(* IEC 61131-3 sources: plc-vscode/tests/st/all/rusty/libs/stdlib/iec61131-st, 25 files *)

(* ---- arithmetic_functions.st ---- *)
(* Definitions of arithmetic functions defined by the IEC61131-3 standard *)

{external}
VAR_GLOBAL
    PI_REAL : REAL;
    PI_LREAL : LREAL;
    FRAC_PI_2_REAL : REAL;
    FRAC_PI_2_LREAL : LREAL;
    FRAC_PI_4_REAL : REAL;
    FRAC_PI_4_LREAL : LREAL;
    E_REAL : REAL;
    E_LREAL : LREAL;
    INF_REAL: REAL;
    INF_LREAL: LREAL;
    NAN_REAL: REAL;
    NAN_LREAL: LREAL;
END_VAR

(********************
*
* This operator returns the value of adding up the operands.
* It overloads the variadic builtin implementation of ADD, which is implemented for ANY_NUM
*
*********************)
FUNCTION ADD < T1: ANY, T2: ANY >: T1
VAR_INPUT
    IN1: T1;
    IN2: T2...;
END_VAR
END_FUNCTION

(********************
*
* This operator produces the multiplication of the operands.
* It overloads the variadic builtin implementation of MUL, which is implemented for ANY_NUM
*
*********************)
FUNCTION MUL < T1: ANY, T2: ANY >: T1
VAR_INPUT
    IN1: T1;
    IN2: T2...;
END_VAR
END_FUNCTION

(* Calculates the square root of a given value *)
{external}
FUNCTION SQRT<T : ANY_REAL> : T
VAR_INPUT
    in : T;
END_VAR
END_FUNCTION

(** Logarithmic functions **)

(* Calculates the natural logarithm of the given value *)
{external}
FUNCTION LN<T : ANY_REAL> : T
VAR_INPUT
    in : T;
END_VAR
END_FUNCTION

(* Calculates the base 10 logarithm of the given value *)
{external}
FUNCTION LOG<T : ANY_REAL> : T
VAR_INPUT
    in : T;
END_VAR
END_FUNCTION

(* Calculates the natural exporenent of the given value *)
{external}
FUNCTION EXP<T : ANY_REAL> : T
VAR_INPUT
    in : T;
END_VAR
END_FUNCTION

(** Trigonometric functions **)

(* Calculates the sine of the given value in radiants *)
{external}
FUNCTION SIN<T : ANY_REAL> : T
VAR_INPUT
    rad : T;
END_VAR
END_FUNCTION

(* Calculates the cosine of the given value in radiants *)
{external}
FUNCTION COS<T : ANY_REAL> : T
VAR_INPUT
    rad : T;
END_VAR
END_FUNCTION

(* Calculates the tangent of the given value in radiants *)
{external}
FUNCTION TAN<T : ANY_REAL> : T
VAR_INPUT
    rad : T;
END_VAR
END_FUNCTION

(* Calculates the arc sine of the given value *)
{external}
FUNCTION ASIN<T : ANY_REAL> : T
VAR_INPUT
    in : T;
END_VAR
END_FUNCTION

(* Calculates the arc cosine of the given value *)
{external}
FUNCTION ACOS<T : ANY_REAL> : T
VAR_INPUT
    in : T;
END_VAR
END_FUNCTION

(* Calculates the arc tangent of the given value *)
{external}
FUNCTION ATAN<T : ANY_REAL> : T
VAR_INPUT
    in : T;
END_VAR
END_FUNCTION

(* Calculate the four quadrant arc tangent of the given values *)
{external}
FUNCTION ATAN2<T : ANY_REAL> : T
VAR_INPUT
    y : T;
    x : T;
END_VAR
END_FUNCTION

{external}
FUNCTION EXPT<T: ANY_REAL, U: ANY_NUM> : T
VAR_INPUT
    in1 : T;
    in2 : U;
END_VAR
END_FUNCTION

{external}
FUNCTION EXPT__REAL__DINT : REAL
VAR_INPUT
    in1 : REAL;
    in2 : DINT;
END_VAR
END_FUNCTION

{external}
FUNCTION EXPT__REAL__REAL : REAL
VAR_INPUT
    in1 : REAL;
    in2 : REAL;
END_VAR
END_FUNCTION

(* LREAL to REAL conversion will happen for the exponent
   This will produce the closest possible REAL value
   On overflow, infinity of the same sign as the input is produced *)
{external}
FUNCTION EXPT__REAL__LREAL : REAL
VAR_INPUT
    in1 : REAL;
    in2 : LREAL;
END_VAR
END_FUNCTION

{external}
FUNCTION EXPT__LREAL__DINT : LREAL
VAR_INPUT
    in1 : LREAL;
    in2 : DINT;
END_VAR
END_FUNCTION

{external}
FUNCTION EXPT__LREAL__REAL : LREAL
VAR_INPUT
    in1 : LREAL;
    in2 : REAL;
END_VAR
END_FUNCTION

{external}
FUNCTION EXPT__LREAL__LREAL : LREAL
VAR_INPUT
    in1 : LREAL;
    in2 : LREAL;
END_VAR
END_FUNCTION

FUNCTION EXPT__REAL__USINT : REAL
VAR_INPUT
    in1 : REAL;
    in2 : USINT;
END_VAR
    EXPT__REAL__USINT := EXPT__REAL__DINT(in1, in2);
END_FUNCTION

FUNCTION EXPT__REAL__UINT : REAL
VAR_INPUT
    in1 : REAL;
    in2 : UINT;
END_VAR
    EXPT__REAL__UINT := EXPT__REAL__DINT(in1, in2);
END_FUNCTION

FUNCTION EXPT__REAL__UDINT : REAL
VAR_INPUT
    in1 : REAL;
    in2 : UDINT;
END_VAR
    EXPT__REAL__UDINT := EXPT__REAL__DINT(in1, in2);
END_FUNCTION

FUNCTION EXPT__REAL__ULINT : REAL
VAR_INPUT
    in1 : REAL;
    in2 : ULINT;
END_VAR
    EXPT__REAL__ULINT := EXPT__REAL__DINT(in1, in2);
END_FUNCTION

FUNCTION EXPT__REAL__SINT : REAL
VAR_INPUT
    in1 : REAL;
    in2 : SINT;
END_VAR
    EXPT__REAL__SINT := EXPT__REAL__DINT(in1, in2);
END_FUNCTION

FUNCTION EXPT__REAL__INT : REAL
VAR_INPUT
    in1 : REAL;
    in2 : INT;
END_VAR
    EXPT__REAL__INT := EXPT__REAL__DINT(in1, in2);
END_FUNCTION

FUNCTION EXPT__REAL__LINT : REAL
VAR_INPUT
    in1 : REAL;
    in2 : LINT;
END_VAR
    EXPT__REAL__LINT := EXPT__REAL__DINT(in1, in2);
END_FUNCTION

FUNCTION EXPT__LREAL__USINT : LREAL
VAR_INPUT
    in1 : LREAL;
    in2 : USINT;
END_VAR
    EXPT__LREAL__USINT := EXPT__LREAL__DINT(in1, in2);
END_FUNCTION

FUNCTION EXPT__LREAL__UINT : LREAL
VAR_INPUT
    in1 : LREAL;
    in2 : UINT;
END_VAR
    EXPT__LREAL__UINT := EXPT__LREAL__DINT(in1, in2);
END_FUNCTION

FUNCTION EXPT__LREAL__UDINT : LREAL
VAR_INPUT
    in1 : LREAL;
    in2 : UDINT;
END_VAR
    EXPT__LREAL__UDINT := EXPT__LREAL__DINT(in1, in2);
END_FUNCTION

FUNCTION EXPT__LREAL__ULINT : LREAL
VAR_INPUT
    in1 : LREAL;
    in2 : ULINT;
END_VAR
    EXPT__LREAL__ULINT := EXPT__LREAL__DINT(in1, in2);
END_FUNCTION

FUNCTION EXPT__LREAL__SINT : LREAL
VAR_INPUT
    in1 : LREAL;
    in2 : SINT;
END_VAR
    EXPT__LREAL__SINT := EXPT__LREAL__DINT(in1, in2);
END_FUNCTION

FUNCTION EXPT__LREAL__INT : LREAL
VAR_INPUT
    in1 : LREAL;
    in2 : INT;
END_VAR
    EXPT__LREAL__INT := EXPT__LREAL__DINT(in1, in2);
END_FUNCTION

FUNCTION EXPT__LREAL__LINT : LREAL
VAR_INPUT
    in1 : LREAL;
    in2 : LINT;
END_VAR
    EXPT__LREAL__LINT := EXPT__LREAL__DINT(in1, in2);
END_FUNCTION

(* ---- string_functions.st ---- *)
VAR_GLOBAL CONSTANT
    __STRING_LENGTH: DINT := 2048;
END_VAR

(* *****************************************************************************
Description: String character length
Input:
    - IN: A character string
Return: String length
***************************************************************************** *)
{external}
FUNCTION LEN < T: ANY_STRING >: DINT
VAR_INPUT {ref}
    IN: T;
END_VAR
END_FUNCTION

(* *****************************************************************************
Description: Left
Input:
    - IN: A character string
    - L: The length of the substring
Return: A substring consisting of the leftmost L characters of IN
***************************************************************************** *)
FUNCTION LEFT < T: ANY_STRING >: T
VAR_INPUT {ref}
    IN: T;
END_VAR
VAR_INPUT
    L: DINT;
END_VAR
END_FUNCTION

{external}
FUNCTION LEFT_EXT < T: ANY_STRING >: DINT
VAR_INPUT {ref}
    IN: T;
END_VAR
VAR_INPUT
    L: DINT;
END_VAR
VAR_IN_OUT
    OUT: T;
END_VAR
END_FUNCTION

FUNCTION LEFT__STRING: STRING[__STRING_LENGTH]
VAR_INPUT {ref}
    IN: STRING[__STRING_LENGTH];
END_VAR
VAR_INPUT
    L: DINT;
END_VAR
    LEFT_EXT(IN, L, LEFT__STRING);
END_FUNCTION

FUNCTION LEFT__WSTRING: WSTRING[__STRING_LENGTH]
VAR_INPUT {ref}
    IN: WSTRING[__STRING_LENGTH];
END_VAR
VAR_INPUT
    L: DINT;
END_VAR
    LEFT_EXT(IN, L, LEFT__WSTRING);
END_FUNCTION

{external}
FUNCTION LEFT_EXT__STRING: DINT
VAR_INPUT {ref}
    IN: STRING[__STRING_LENGTH];
END_VAR
VAR_INPUT
    L: DINT;
END_VAR
VAR_IN_OUT
    OUT: STRING[__STRING_LENGTH];
END_VAR
END_FUNCTION

{external}
FUNCTION LEFT_EXT__WSTRING: DINT
VAR_INPUT {ref}
    IN: WSTRING[__STRING_LENGTH];
END_VAR
VAR_INPUT
    L: DINT;
END_VAR
VAR_IN_OUT
    OUT: WSTRING[__STRING_LENGTH];
END_VAR
END_FUNCTION

(* *****************************************************************************
Description: Right
Input:
    - IN: A character string
    - L: The length of the substring
Return: A substring consisting of the rightmost L characters of IN
***************************************************************************** *)
FUNCTION RIGHT < T: ANY_STRING >: T
VAR_INPUT {ref}
    IN: T;
END_VAR
VAR_INPUT
    L: DINT;
END_VAR
END_FUNCTION

{external}
FUNCTION RIGHT_EXT < T: ANY_STRING >: DINT
VAR_INPUT {ref}
    IN: T;
END_VAR
VAR_INPUT
    L: DINT;
END_VAR
VAR_IN_OUT
    OUT: T;
END_VAR
END_FUNCTION

FUNCTION RIGHT__STRING: STRING[__STRING_LENGTH]
VAR_INPUT {ref}
    IN: STRING[__STRING_LENGTH];
END_VAR
VAR_INPUT
    L: DINT;
END_VAR
    RIGHT_EXT(IN, L, RIGHT__STRING);
END_FUNCTION

FUNCTION RIGHT__WSTRING: WSTRING[__STRING_LENGTH]
VAR_INPUT {ref}
    IN: WSTRING[__STRING_LENGTH];
END_VAR
VAR_INPUT
    L: DINT;
END_VAR
    RIGHT_EXT(IN, L, RIGHT__WSTRING);
END_FUNCTION

{external}
FUNCTION RIGHT_EXT__STRING: DINT
VAR_INPUT {ref}
    IN: STRING[__STRING_LENGTH];
END_VAR
VAR_INPUT
    L: DINT;
END_VAR
VAR_IN_OUT
    OUT: STRING[__STRING_LENGTH];
END_VAR
END_FUNCTION

{external}
FUNCTION RIGHT_EXT__WSTRING: DINT
VAR_INPUT {ref}
    IN: WSTRING[__STRING_LENGTH];
END_VAR
VAR_INPUT
    L: DINT;
END_VAR
VAR_IN_OUT
    OUT: WSTRING[__STRING_LENGTH];
END_VAR
END_FUNCTION

(* *****************************************************************************
Description: Middle
Input:
    - IN: A character string
    - L: The length of the substring
    - P: The starting index position
Return:
    A substring that contains L characters starting
    from position P in a string.
***************************************************************************** *)
FUNCTION MID < T: ANY_STRING >: T
VAR_INPUT {ref}
    IN: T;
END_VAR
VAR_INPUT
    L: DINT;
    P: DINT;
END_VAR
END_FUNCTION

{external}
FUNCTION MID_EXT < T: ANY_STRING >: DINT
VAR_INPUT {ref}
    IN: T;
END_VAR
VAR_INPUT
    L: DINT;
    P: DINT;
END_VAR
VAR_IN_OUT
    OUT: T;
END_VAR
END_FUNCTION

FUNCTION MID__STRING: STRING[__STRING_LENGTH]
VAR_INPUT {ref}
    IN: STRING[__STRING_LENGTH];
END_VAR
VAR_INPUT
    L: DINT;
    P: DINT;
END_VAR
    MID_EXT(IN, L, P, MID__STRING);
END_FUNCTION

FUNCTION MID__WSTRING: WSTRING[__STRING_LENGTH]
VAR_INPUT {ref}
    IN: WSTRING[__STRING_LENGTH];
END_VAR
VAR_INPUT
    L: DINT;
    P: DINT;
END_VAR
    MID_EXT(IN, L, P, MID__WSTRING);
END_FUNCTION

{external}
FUNCTION MID_EXT__STRING: DINT
VAR_INPUT {ref}
    IN: STRING[__STRING_LENGTH];
END_VAR
VAR_INPUT
    L: DINT;
    P: DINT;
END_VAR
VAR_IN_OUT
    OUT: STRING[__STRING_LENGTH];
END_VAR
END_FUNCTION

{external}
FUNCTION MID_EXT__WSTRING: DINT
VAR_INPUT {ref}
    IN: WSTRING[__STRING_LENGTH];
END_VAR
VAR_INPUT
    L: DINT;
    P: DINT;
END_VAR
VAR_IN_OUT
    OUT: WSTRING[__STRING_LENGTH];
END_VAR
END_FUNCTION

(* *****************************************************************************
Description: Extensible concatenation
Input:
    - IN: Two or more comma-separated strings
Return:
    A string combining all given input strings in the same order
    as the given string parameters.
***************************************************************************** *)
{external}
FUNCTION CONCAT__STRING: STRING[2048]
VAR_INPUT {ref}
    args: {sized} STRING...;
END_VAR
END_FUNCTION

{external}
FUNCTION CONCAT__WSTRING: WSTRING[2048]
VAR_INPUT {ref}
    args: {sized} WSTRING...;
END_VAR
END_FUNCTION

FUNCTION CONCAT < T: ANY_STRING >: T
VAR_INPUT {ref}
    args: {sized} T...;
END_VAR
END_FUNCTION

{external}
FUNCTION CONCAT_EXT < T: ANY_STRING >: DINT
VAR_IN_OUT
    OUT: T;
END_VAR
VAR_INPUT {ref}
    args: {sized} T...;
END_VAR
END_FUNCTION

(* *****************************************************************************
Description: Insert
Input:
    IN1: The string to insert into
    IN2: The string to insert
    P: The position at which to insert
Return:
    A string consisting of IN2 inserted at position P into string IN1
***************************************************************************** *)
FUNCTION INSERT < T: ANY_STRING >: T
VAR_INPUT {ref}
    IN1: T;
    IN2: T;
END_VAR
VAR_INPUT
    P: DINT;
END_VAR
END_FUNCTION

{external}
FUNCTION INSERT_EXT < T: ANY_STRING >: DINT
VAR_INPUT {ref}
    IN1: T;
    IN2: T;
END_VAR
VAR_INPUT
    P: DINT;
END_VAR
VAR_IN_OUT
    OUT: T;
END_VAR
END_FUNCTION

FUNCTION INSERT__STRING: STRING[__STRING_LENGTH]
VAR_INPUT {ref}
    IN1: STRING[__STRING_LENGTH];
    IN2: STRING[__STRING_LENGTH];
END_VAR
VAR_INPUT
    P: DINT;
END_VAR
    INSERT_EXT(IN1, IN2, P, INSERT__STRING);
END_FUNCTION

FUNCTION INSERT__WSTRING: WSTRING[__STRING_LENGTH]
VAR_INPUT {ref}
    IN1: WSTRING[__STRING_LENGTH];
    IN2: WSTRING[__STRING_LENGTH];
END_VAR
VAR_INPUT
    P: DINT;
END_VAR
    INSERT_EXT(IN1, IN2, P, INSERT__WSTRING);
END_FUNCTION

{external}
FUNCTION INSERT_EXT__STRING: DINT
VAR_INPUT {ref}
    IN1: STRING[__STRING_LENGTH];
    IN2: STRING[__STRING_LENGTH];
END_VAR
VAR_INPUT
    P: DINT;
END_VAR
VAR_IN_OUT
    OUT: STRING[__STRING_LENGTH];
END_VAR
END_FUNCTION

{external}
FUNCTION INSERT_EXT__WSTRING: DINT
VAR_INPUT {ref}
    IN1: WSTRING[__STRING_LENGTH];
    IN2: WSTRING[__STRING_LENGTH];
END_VAR
VAR_INPUT
    P: DINT;
END_VAR
VAR_IN_OUT
    OUT: WSTRING[__STRING_LENGTH];
END_VAR
END_FUNCTION

(* *****************************************************************************
Description: Delete
Input:
    IN: The string to delete characters from
    L: The amount of characters to delete
    P: The position at which to start deleting
Return: A new string with L characters deleted from P onwards
***************************************************************************** *)
FUNCTION DELETE < T: ANY_STRING >: T
VAR_INPUT {ref}
    IN: T;
END_VAR
VAR_INPUT
    L: DINT;
    P: DINT;
END_VAR
END_FUNCTION

{external}
FUNCTION DELETE_EXT < T: ANY_STRING >: DINT
VAR_INPUT {ref}
    IN: T;
END_VAR
VAR_INPUT
    L: DINT;
    P: DINT;
END_VAR
VAR_IN_OUT
    OUT: T;
END_VAR
END_FUNCTION

FUNCTION DELETE__STRING: STRING[__STRING_LENGTH]
VAR_INPUT {ref}
    IN: STRING[__STRING_LENGTH];
END_VAR
VAR_INPUT
    L: DINT;
    P: DINT;
END_VAR
    DELETE_EXT(IN, L, P, DELETE__STRING);
END_FUNCTION

FUNCTION DELETE__WSTRING: WSTRING[__STRING_LENGTH]
VAR_INPUT {ref}
    IN: WSTRING[__STRING_LENGTH];
END_VAR
VAR_INPUT
    L: DINT;
    P: DINT;
END_VAR
    DELETE_EXT(IN, L, P, DELETE__WSTRING);
END_FUNCTION

{external}
FUNCTION DELETE_EXT__STRING: DINT
VAR_INPUT {ref}
    IN: STRING[__STRING_LENGTH];
END_VAR
VAR_INPUT
    L: DINT;
    P: DINT;
END_VAR
VAR_IN_OUT
    OUT: STRING[__STRING_LENGTH];
END_VAR
END_FUNCTION

{external}
FUNCTION DELETE_EXT__WSTRING: DINT
VAR_INPUT {ref}
    IN: WSTRING[__STRING_LENGTH];
END_VAR
VAR_INPUT
    L: DINT;
    P: DINT;
END_VAR
VAR_IN_OUT
    OUT: WSTRING[__STRING_LENGTH];
END_VAR
END_FUNCTION
(* *****************************************************************************
Description: Replace
Input:
    IN1: The string to replace characters from
    IN2: The replacement string to be inserted
    L: The amount of characters to delete
    P: The position at which to start deleting
Return: A new string which has L characters replaced by IN2 from position P onwards
***************************************************************************** *)
FUNCTION REPLACE < T: ANY_STRING >: T
VAR_INPUT {ref}
    IN1: T;
    IN2: T;
END_VAR
VAR_INPUT
    L: DINT;
    P: DINT;
END_VAR
END_FUNCTION

{external}
FUNCTION REPLACE_EXT < T: ANY_STRING >: DINT
VAR_INPUT {ref}
    IN1: T;
    IN2: T;
END_VAR
VAR_INPUT
    L: DINT;
    P: DINT;
END_VAR
VAR_IN_OUT
    OUT: T;
END_VAR
END_FUNCTION

FUNCTION REPLACE__STRING: STRING[__STRING_LENGTH]
VAR_INPUT {ref}
    IN1: STRING[__STRING_LENGTH];
    IN2: STRING[__STRING_LENGTH];
END_VAR
VAR_INPUT
    L: DINT;
    P: DINT;
END_VAR
    REPLACE_EXT(IN1, IN2, L, P, REPLACE__STRING);
END_FUNCTION

FUNCTION REPLACE__WSTRING: WSTRING[__STRING_LENGTH]
VAR_INPUT {ref}
    IN1: WSTRING[__STRING_LENGTH];
    IN2: WSTRING[__STRING_LENGTH];
END_VAR
VAR_INPUT
    L: DINT;
    P: DINT;
END_VAR
    REPLACE_EXT(IN1, IN2, L, P, REPLACE__WSTRING);
END_FUNCTION

{external}
FUNCTION REPLACE_EXT__STRING: DINT
VAR_INPUT {ref}
    IN1: STRING[__STRING_LENGTH];
    IN2: STRING[__STRING_LENGTH];
END_VAR
VAR_INPUT
    L: DINT;
    P: DINT;
END_VAR
VAR_IN_OUT
    OUT: STRING[__STRING_LENGTH];
END_VAR
END_FUNCTION

{external}
FUNCTION REPLACE_EXT__WSTRING: DINT
VAR_INPUT {ref}
    IN1: WSTRING[__STRING_LENGTH];
    IN2: WSTRING[__STRING_LENGTH];
END_VAR
VAR_INPUT
    L: DINT;
    P: DINT;
END_VAR
VAR_IN_OUT
    OUT: WSTRING[__STRING_LENGTH];
END_VAR
END_FUNCTION

(* *****************************************************************************
Description: Find
Input:
    IN1: The string in which to search in
    IN2: The substring to search for
Return: The character index of the first match. 0 if there are no matches.
***************************************************************************** *)
{external}
FUNCTION FIND < T: ANY_STRING >: DINT
VAR_INPUT {ref}
    IN1: T;
    IN2: T;
END_VAR
END_FUNCTION

(* *****************************************************************************
Description: Decreasing sequence
Input: The strings to compare, in order. ((IN1>IN2) & (IN2>IN3) & .. & (INn-1>INn))
Return:
    TRUE if codepoints are in decreasing order (alphabetical order: ZYX > YXW > XWV ..)
    FALSE otherwise
***************************************************************************** *)
// passing strings by ref causes an error/warning. code still compiles and works correctly
FUNCTION STRING_GREATER: BOOL
VAR_INPUT
    a, b: STRING;
END_VAR
    STRING_GREATER := __STRING_GREATER(a, b);
END_FUNCTION

FUNCTION WSTRING_GREATER: BOOL
VAR_INPUT
    a, b: WSTRING;
END_VAR
    WSTRING_GREATER := __WSTRING_GREATER(a, b);
END_FUNCTION

(* *****************************************************************************
Description: Equality
Input: The strings to compare, in order. ((IN1=IN2) & (IN2=IN3) & .. & (INn-1=INn))
Return:
    TRUE if codepoints are equal to each other
    FALSE otherwise.
***************************************************************************** *)
FUNCTION STRING_EQUAL: BOOL
VAR_INPUT
    a, b: STRING;
END_VAR
    STRING_EQUAL := __STRING_EQUAL(a, b);
END_FUNCTION

FUNCTION WSTRING_EQUAL: BOOL
VAR_INPUT
    a, b: WSTRING;
END_VAR
    WSTRING_EQUAL := __WSTRING_EQUAL(a, b);
END_FUNCTION

(* *****************************************************************************
Description: Increasing sequence
Input: The strings to compare, in order. ((IN1<IN2) & (IN2<IN3) & .. & (INn-1<INn))
Return:
    TRUE if codepoints are in increasing order (alphabetical order: ABC < BCD < CDE ..)
    FALSE otherwise
***************************************************************************** *)
FUNCTION STRING_LESS: BOOL
VAR_INPUT
    a, b: STRING;
END_VAR
    STRING_LESS := __STRING_LESS(a, b);
END_FUNCTION

FUNCTION WSTRING_LESS: BOOL
VAR_INPUT
    a, b: WSTRING;
END_VAR
    WSTRING_LESS := __WSTRING_LESS(a, b);
END_FUNCTION

// internal functions
{external}
FUNCTION __STRING_GREATER: BOOL
VAR_INPUT {ref}
    IN: {sized} STRING...;
END_VAR
END_FUNCTION

{external}
FUNCTION __STRING_EQUAL: BOOL
VAR_INPUT {ref}
    IN: {sized} STRING...;
END_VAR
END_FUNCTION

{external}
FUNCTION __STRING_LESS: BOOL
VAR_INPUT {ref}
    IN: {sized} STRING...;
END_VAR
END_FUNCTION

{external}
FUNCTION __WSTRING_GREATER: BOOL
VAR_INPUT {ref}
    IN: {sized} WSTRING...;
END_VAR
END_FUNCTION

{external}
FUNCTION __WSTRING_EQUAL: BOOL
VAR_INPUT {ref}
    IN: {sized} WSTRING...;
END_VAR
END_FUNCTION

{external}
FUNCTION __WSTRING_LESS: BOOL
VAR_INPUT {ref}
    IN: {sized} WSTRING...;
END_VAR
END_FUNCTION

(* ---- bit_conversion.st ---- *)
(********************
*
* Converts LWORD to DWORD
*
*********************)
FUNCTION LWORD_TO_DWORD : DWORD
VAR_INPUT
    in : LWORD;
END_VAR
    LWORD_TO_DWORD := in;
END_FUNCTION

(********************
*
* Converts LWORD to WORD
*
*********************)
FUNCTION LWORD_TO_WORD : WORD
VAR_INPUT
    in : LWORD;
END_VAR
    LWORD_TO_WORD := in;
END_FUNCTION

(********************
*
* Converts LWORD to BYTE
*
*********************)
FUNCTION LWORD_TO_BYTE : BYTE
VAR_INPUT
    in : LWORD;
END_VAR
    LWORD_TO_BYTE := in;
END_FUNCTION

(********************
*
* Converts LWORD to BOOL
*
*********************)
FUNCTION LWORD_TO_BOOL : BOOL
VAR_INPUT
    in : LWORD;
END_VAR
    LWORD_TO_BOOL := in.0;
END_FUNCTION

(********************
*
* Converts DWORD to LWORD
*
*********************)
FUNCTION DWORD_TO_LWORD : LWORD
VAR_INPUT
    in : DWORD;
END_VAR
    DWORD_TO_LWORD := in;
END_FUNCTION

(********************
*
* Converts DWORD to WORD
*
*********************)
FUNCTION DWORD_TO_WORD : WORD
VAR_INPUT
    in : DWORD;
END_VAR
    DWORD_TO_WORD := in;
END_FUNCTION

(********************
*
* Converts DWORD to BYTE
*
*********************)
FUNCTION DWORD_TO_BYTE : BYTE
VAR_INPUT
    in : DWORD;
END_VAR
    DWORD_TO_BYTE := in;
END_FUNCTION

(********************
*
* Converts DWORD to BOOL
*
*********************)
FUNCTION DWORD_TO_BOOL : BOOL
VAR_INPUT
    in : DWORD;
END_VAR
    DWORD_TO_BOOL := in.0;
END_FUNCTION

(********************
*
* Converts WORD to LWORD
*
*********************)
FUNCTION WORD_TO_LWORD : LWORD
VAR_INPUT
    in : WORD;
END_VAR
    WORD_TO_LWORD := in;
END_FUNCTION

(********************
*
* Converts WORD to DWORD
*
*********************)
FUNCTION WORD_TO_DWORD : DWORD
VAR_INPUT
    in : WORD;
END_VAR
    WORD_TO_DWORD := in;
END_FUNCTION

(********************
*
* Converts WORD to BYTE
*
*********************)
FUNCTION WORD_TO_BYTE : BYTE
VAR_INPUT
    in : WORD;
END_VAR
    WORD_TO_BYTE := in;
END_FUNCTION

(********************
*
* Converts WORD to BOOL
*
*********************)
FUNCTION WORD_TO_BOOL : BOOL
VAR_INPUT
    in : WORD;
END_VAR
    WORD_TO_BOOL := in.0;
END_FUNCTION

(********************
*
* Converts BYTE to LWORD
*
*********************)
FUNCTION BYTE_TO_LWORD : LWORD
VAR_INPUT
    in : BYTE;
END_VAR
    BYTE_TO_LWORD := in;
END_FUNCTION

(********************
*
* Converts BYTE to DWORD
*
*********************)
FUNCTION BYTE_TO_DWORD : DWORD
VAR_INPUT
    in : BYTE;
END_VAR
    BYTE_TO_DWORD := in;
END_FUNCTION

(********************
*
* Converts BYTE to WORD
*
*********************)
FUNCTION BYTE_TO_WORD : WORD
VAR_INPUT
    in : BYTE;
END_VAR
    BYTE_TO_WORD := in;
END_FUNCTION

(********************
*
* Converts BYTE to BOOL
*
*********************)
FUNCTION BYTE_TO_BOOL : BOOL
VAR_INPUT
    in : BYTE;
END_VAR
    BYTE_TO_BOOL := in.0;
END_FUNCTION

(********************
*
* Converts BYTE to CHAR
*
*********************)
FUNCTION BYTE_TO_CHAR : CHAR
VAR_INPUT
    in : BYTE;
END_VAR
VAR
    ptr : REF_TO CHAR;
END_VAR
    ptr := REF(in);
    BYTE_TO_CHAR := ptr^;
END_FUNCTION

(********************
*
* Converts BOOL to LWORD
*
*********************)
FUNCTION BOOL_TO_LWORD : LWORD
VAR_INPUT
    in : BOOL;
END_VAR
    IF in <> 0 THEN
        BOOL_TO_LWORD := 1;
    ELSE
        BOOL_TO_LWORD := 0;
    END_IF;
END_FUNCTION

(********************
*
* Converts BOOL to DWORD
*
*********************)
FUNCTION BOOL_TO_DWORD : DWORD
VAR_INPUT
    in : BOOL;
END_VAR
    IF in <> 0 THEN
        BOOL_TO_DWORD := 1;
    ELSE
        BOOL_TO_DWORD := 0;
    END_IF;
END_FUNCTION

(********************
*
* Converts BOOL to WORD
*
*********************)
FUNCTION BOOL_TO_WORD : WORD
VAR_INPUT
    in : BOOL;
END_VAR
    IF in <> 0 THEN
        BOOL_TO_WORD := 1;
    ELSE
        BOOL_TO_WORD := 0;
    END_IF;
END_FUNCTION

(********************
*
* Converts BOOL to BYTE
*
*********************)
FUNCTION BOOL_TO_BYTE : BYTE
VAR_INPUT
    in : BOOL;
END_VAR
    IF in <> 0 THEN
        BOOL_TO_BYTE := 1;
    ELSE
        BOOL_TO_BYTE := 0;
    END_IF;
END_FUNCTION

(********************
*
* Converts CHAR to BYTE
*
*********************)
FUNCTION CHAR_TO_BYTE : BYTE
VAR_INPUT
    in : CHAR;
END_VAR
VAR
    ptr : REF_TO BYTE;
END_VAR
    ptr := REF(in);
    CHAR_TO_BYTE := ptr^;
END_FUNCTION

(********************
*
* Converts WCHAR to BYTE
*
*********************)
FUNCTION WCHAR_TO_BYTE : BYTE
VAR_INPUT
    in : WCHAR;
END_VAR
VAR
    ptr : REF_TO BYTE;
END_VAR
    ptr := REF(in);
    WCHAR_TO_BYTE := ptr^;
END_FUNCTION

(********************
*
* Converts CHAR to WORD
*
*********************)
FUNCTION CHAR_TO_WORD : WORD
VAR_INPUT
    in : CHAR;
END_VAR
    CHAR_TO_WORD := CHAR_TO_BYTE(in);
END_FUNCTION

(********************
*
* Converts CHAR to DWORD
*
*********************)
FUNCTION CHAR_TO_DWORD : DWORD
VAR_INPUT
    in : CHAR;
END_VAR
    CHAR_TO_DWORD := CHAR_TO_BYTE(in);
END_FUNCTION

(********************
*
* Converts CHAR to LWORD
*
*********************)
FUNCTION CHAR_TO_LWORD : LWORD
VAR_INPUT
    in : CHAR;
END_VAR
    CHAR_TO_LWORD := CHAR_TO_BYTE(in);
END_FUNCTION

(********************
*
* Converts WCHAR to WORD
*
*********************)
FUNCTION WCHAR_TO_WORD : WORD
VAR_INPUT
    in : WCHAR;
END_VAR
VAR
    ptr : REF_TO WORD;
END_VAR
    ptr := REF(in);
    WCHAR_TO_WORD := ptr^;
END_FUNCTION

(********************
*
* Converts WCHAR to DWORD
*
*********************)
FUNCTION WCHAR_TO_DWORD : DWORD
VAR_INPUT
    in : WCHAR;
END_VAR
    WCHAR_TO_DWORD := WCHAR_TO_WORD(in);
END_FUNCTION

(********************
*
* Converts WCHAR to LWORD
*
*********************)
FUNCTION WCHAR_TO_LWORD : LWORD
VAR_INPUT
    in : WCHAR;
END_VAR
    WCHAR_TO_LWORD := WCHAR_TO_WORD(in);
END_FUNCTION

(* ---- bit_num_conversion.st ---- *)
(********************
*
* Converts LWORD to LREAL
*
*********************)
{external}
FUNCTION LWORD_TO_LREAL : LREAL
VAR_INPUT
    in : LWORD;
END_VAR
END_FUNCTION

(********************
*
* Converts LWORD to LINT
*
*********************)
FUNCTION LWORD_TO_LINT : LINT
VAR_INPUT
    in : LWORD;
END_VAR
    LWORD_TO_LINT := in;
END_FUNCTION

(********************
*
* Converts LWORD to DINT
*
*********************)
FUNCTION LWORD_TO_DINT : DINT
VAR_INPUT
    in : LWORD;
END_VAR
    LWORD_TO_DINT := in;
END_FUNCTION

(********************
*
* Converts LWORD to INT
*
*********************)
FUNCTION LWORD_TO_INT : INT
VAR_INPUT
    in : LWORD;
END_VAR
    LWORD_TO_INT := in;
END_FUNCTION

(********************
*
* Converts LWORD to SINT
*
*********************)
FUNCTION LWORD_TO_SINT : SINT
VAR_INPUT
    in : LWORD;
END_VAR
    LWORD_TO_SINT := in;
END_FUNCTION

(********************
*
* Converts LWORD to ULINT
*
*********************)
FUNCTION LWORD_TO_ULINT : ULINT
VAR_INPUT
    in : LWORD;
END_VAR
    LWORD_TO_ULINT := in;
END_FUNCTION

(********************
*
* Converts LWORD to UDINT
*
*********************)
FUNCTION LWORD_TO_UDINT : UDINT
VAR_INPUT
    in : LWORD;
END_VAR
    LWORD_TO_UDINT := in;
END_FUNCTION

(********************
*
* Converts LWORD to UINT
*
*********************)
FUNCTION LWORD_TO_UINT : UINT
VAR_INPUT
    in : LWORD;
END_VAR
    LWORD_TO_UINT := in;
END_FUNCTION

(********************
*
* Converts LWORD to USINT
*
*********************)
FUNCTION LWORD_TO_USINT : USINT
VAR_INPUT
    in : LWORD;
END_VAR
    LWORD_TO_USINT := in;
END_FUNCTION

(********************
*
* Converts DWORD to REAL
*
*********************)
{external}
FUNCTION DWORD_TO_REAL : REAL
VAR_INPUT
    in : DWORD;
END_VAR
END_FUNCTION

(********************
*
* Converts DWORD to LINT
*
*********************)
FUNCTION DWORD_TO_LINT : LINT
VAR_INPUT
    in : DWORD;
END_VAR
    DWORD_TO_LINT := in;
END_FUNCTION

(********************
*
* Converts DWORD to DINT
*
*********************)
FUNCTION DWORD_TO_DINT : DINT
VAR_INPUT
    in : DWORD;
END_VAR
    DWORD_TO_DINT := in;
END_FUNCTION

(********************
*
* Converts DWORD to INT
*
*********************)
FUNCTION DWORD_TO_INT : INT
VAR_INPUT
    in : DWORD;
END_VAR
    DWORD_TO_INT := in;
END_FUNCTION

(********************
*
* Converts DWORD to SINT
*
*********************)
FUNCTION DWORD_TO_SINT : SINT
VAR_INPUT
    in : DWORD;
END_VAR
    DWORD_TO_SINT := in;
END_FUNCTION

(********************
*
* Converts DWORD to ULINT
*
*********************)
FUNCTION DWORD_TO_ULINT : ULINT
VAR_INPUT
    in : DWORD;
END_VAR
    DWORD_TO_ULINT := in;
END_FUNCTION

(********************
*
* Converts DWORD to UDINT
*
*********************)
FUNCTION DWORD_TO_UDINT : UDINT
VAR_INPUT
    in : DWORD;
END_VAR
    DWORD_TO_UDINT := in;
END_FUNCTION

(********************
*
* Converts DWORD to UINT
*
*********************)
FUNCTION DWORD_TO_UINT : UINT
VAR_INPUT
    in : DWORD;
END_VAR
    DWORD_TO_UINT := in;
END_FUNCTION

(********************
*
* Converts DWORD to USINT
*
*********************)
FUNCTION DWORD_TO_USINT : USINT
VAR_INPUT
    in : DWORD;
END_VAR
    DWORD_TO_USINT := in;
END_FUNCTION

(********************
*
* Converts WORD to LINT
*
*********************)
FUNCTION WORD_TO_LINT : LINT
VAR_INPUT
    in : WORD;
END_VAR
    WORD_TO_LINT := in;
END_FUNCTION

(********************
*
* Converts WORD to DINT
*
*********************)
FUNCTION WORD_TO_DINT : DINT
VAR_INPUT
    in : WORD;
END_VAR
    WORD_TO_DINT := in;
END_FUNCTION

(********************
*
* Converts WORD to INT
*
*********************)
FUNCTION WORD_TO_INT : INT
VAR_INPUT
    in : WORD;
END_VAR
    WORD_TO_INT := in;
END_FUNCTION

(********************
*
* Converts WORD to SINT
*
*********************)
FUNCTION WORD_TO_SINT : SINT
VAR_INPUT
    in : WORD;
END_VAR
    WORD_TO_SINT := in;
END_FUNCTION

(********************
*
* Converts WORD to ULINT
*
*********************)
FUNCTION WORD_TO_ULINT : ULINT
VAR_INPUT
    in : WORD;
END_VAR
    WORD_TO_ULINT := in;
END_FUNCTION

(********************
*
* Converts WORD to UDINT
*
*********************)
FUNCTION WORD_TO_UDINT : UDINT
VAR_INPUT
    in : WORD;
END_VAR
    WORD_TO_UDINT := in;
END_FUNCTION

(********************
*
* Converts WORD to UINT
*
*********************)
FUNCTION WORD_TO_UINT : UINT
VAR_INPUT
    in : WORD;
END_VAR
    WORD_TO_UINT := in;
END_FUNCTION

(********************
*
* Converts WORD to USINT
*
*********************)
FUNCTION WORD_TO_USINT : USINT
VAR_INPUT
    in : WORD;
END_VAR
    WORD_TO_USINT := in;
END_FUNCTION

(********************
*
* Converts BYTE to LINT
*
*********************)
FUNCTION BYTE_TO_LINT : LINT
VAR_INPUT
    in : BYTE;
END_VAR
    BYTE_TO_LINT := in;
END_FUNCTION

(********************
*
* Converts BYTE to DINT
*
*********************)
FUNCTION BYTE_TO_DINT : DINT
VAR_INPUT
    in : BYTE;
END_VAR
    BYTE_TO_DINT := in;
END_FUNCTION

(********************
*
* Converts BYTE to INT
*
*********************)
FUNCTION BYTE_TO_INT : INT
VAR_INPUT
    in : BYTE;
END_VAR
    BYTE_TO_INT := in;
END_FUNCTION

(********************
*
* Converts BYTE to SINT
*
*********************)
FUNCTION BYTE_TO_SINT : SINT
VAR_INPUT
    in : BYTE;
END_VAR
    BYTE_TO_SINT := in;
END_FUNCTION

(********************
*
* Converts BYTE to ULINT
*
*********************)
FUNCTION BYTE_TO_ULINT : ULINT
VAR_INPUT
    in : BYTE;
END_VAR
    BYTE_TO_ULINT := in;
END_FUNCTION

(********************
*
* Converts BYTE to UDINT
*
*********************)
FUNCTION BYTE_TO_UDINT : UDINT
VAR_INPUT
    in : BYTE;
END_VAR
    BYTE_TO_UDINT := in;
END_FUNCTION

(********************
*
* Converts BYTE to UINT
*
*********************)
FUNCTION BYTE_TO_UINT : UINT
VAR_INPUT
    in : BYTE;
END_VAR
    BYTE_TO_UINT := in;
END_FUNCTION

(********************
*
* Converts BYTE to USINT
*
*********************)
FUNCTION BYTE_TO_USINT : USINT
VAR_INPUT
    in : BYTE;
END_VAR
    BYTE_TO_USINT := in;
END_FUNCTION

(********************
*
* Converts BOOL to LINT
*
*********************)
FUNCTION BOOL_TO_LINT : LINT
VAR_INPUT
    in : BOOL;
END_VAR
    BOOL_TO_LINT := in;
END_FUNCTION

(********************
*
* Converts BOOL to DINT
*
*********************)
FUNCTION BOOL_TO_DINT : DINT
VAR_INPUT
    in : BOOL;
END_VAR
    BOOL_TO_DINT := in;
END_FUNCTION

(********************
*
* Converts BOOL to INT
*
*********************)
FUNCTION BOOL_TO_INT : INT
VAR_INPUT
    in : BOOL;
END_VAR
    BOOL_TO_INT := in;
END_FUNCTION

(********************
*
* Converts BOOL to SINT
*
*********************)
FUNCTION BOOL_TO_SINT : SINT
VAR_INPUT
    in : BOOL;
END_VAR
    BOOL_TO_SINT := in;
END_FUNCTION

(********************
*
* Converts BOOL to ULINT
*
*********************)
FUNCTION BOOL_TO_ULINT : ULINT
VAR_INPUT
    in : BOOL;
END_VAR
    BOOL_TO_ULINT := in;
END_FUNCTION

(********************
*
* Converts BOOL to UDINT
*
*********************)
FUNCTION BOOL_TO_UDINT : UDINT
VAR_INPUT
    in : BOOL;
END_VAR
    BOOL_TO_UDINT := in;
END_FUNCTION

(********************
*
* Converts BOOL to UINT
*
*********************)
FUNCTION BOOL_TO_UINT : UINT
VAR_INPUT
    in : BOOL;
END_VAR
    BOOL_TO_UINT := in;
END_FUNCTION

(********************
*
* Converts BOOL to USINT
*
*********************)
FUNCTION BOOL_TO_USINT : USINT
VAR_INPUT
    in : BOOL;
END_VAR
    BOOL_TO_USINT := in;
END_FUNCTION

(********************
*
* Converts LREAL to LWORD
*
*********************)
{external}
FUNCTION LREAL_TO_LWORD : LWORD
VAR_INPUT
    in : LREAL;
END_VAR
END_FUNCTION

(********************
*
* Converts REAL to DWORD
*
*********************)
{external}
FUNCTION REAL_TO_DWORD : DWORD
VAR_INPUT
    in : REAL;
END_VAR
END_FUNCTION

(********************
*
* Converts LINT to LWORD
*
*********************)
FUNCTION LINT_TO_LWORD : LWORD
VAR_INPUT
    in : LINT;
END_VAR
    LINT_TO_LWORD := in;
END_FUNCTION

(********************
*
* Converts LINT to DWORD
*
*********************)
FUNCTION LINT_TO_DWORD : DWORD
VAR_INPUT
    in : LINT;
END_VAR
    LINT_TO_DWORD := in;
END_FUNCTION

(********************
*
* Converts LINT to WORD
*
*********************)
FUNCTION LINT_TO_WORD : WORD
VAR_INPUT
    in : LINT;
END_VAR
    LINT_TO_WORD := in;
END_FUNCTION

(********************
*
* Converts LINT to BYTE
*
*********************)
FUNCTION LINT_TO_BYTE : BYTE
VAR_INPUT
    in : LINT;
END_VAR
    LINT_TO_BYTE := in;
END_FUNCTION

(********************
*
* Converts DINT to LWORD
*
*********************)
FUNCTION DINT_TO_LWORD : LWORD
VAR_INPUT
    in : DINT;
END_VAR
    DINT_TO_LWORD := in;
END_FUNCTION

(********************
*
* Converts DINT to DWORD
*
*********************)
FUNCTION DINT_TO_DWORD : DWORD
VAR_INPUT
    in : DINT;
END_VAR
    DINT_TO_DWORD := in;
END_FUNCTION

(********************
*
* Converts DINT to WORD
*
*********************)
FUNCTION DINT_TO_WORD : WORD
VAR_INPUT
    in : DINT;
END_VAR
    DINT_TO_WORD := in;
END_FUNCTION

(********************
*
* Converts DINT to BYTE
*
*********************)
FUNCTION DINT_TO_BYTE : BYTE
VAR_INPUT
    in : DINT;
END_VAR
    DINT_TO_BYTE := in;
END_FUNCTION

(********************
*
* Converts INT to LWORD
*
*********************)
FUNCTION INT_TO_LWORD : LWORD
VAR_INPUT
    in : INT;
END_VAR
    INT_TO_LWORD := in;
END_FUNCTION

(********************
*
* Converts INT to DWORD
*
*********************)
FUNCTION INT_TO_DWORD : DWORD
VAR_INPUT
    in : INT;
END_VAR
    INT_TO_DWORD := in;
END_FUNCTION

(********************
*
* Converts INT to WORD
*
*********************)
FUNCTION INT_TO_WORD : WORD
VAR_INPUT
    in : INT;
END_VAR
    INT_TO_WORD := in;
END_FUNCTION

(********************
*
* Converts INT to BYTE
*
*********************)
FUNCTION INT_TO_BYTE : BYTE
VAR_INPUT
    in : INT;
END_VAR
    INT_TO_BYTE := in;
END_FUNCTION

(********************
*
* Converts SINT to LWORD
*
*********************)
FUNCTION SINT_TO_LWORD : LWORD
VAR_INPUT
    in : SINT;
END_VAR
    SINT_TO_LWORD := in;
END_FUNCTION

(********************
*
* Converts SINT to DWORD
*
*********************)
FUNCTION SINT_TO_DWORD : DWORD
VAR_INPUT
    in : SINT;
END_VAR
    SINT_TO_DWORD := in;
END_FUNCTION

(********************
*
* Converts SINT to WORD
*
*********************)
FUNCTION SINT_TO_WORD : WORD
VAR_INPUT
    in : SINT;
END_VAR
    SINT_TO_WORD := in;
END_FUNCTION

(********************
*
* Converts SINT to BYTE
*
*********************)
FUNCTION SINT_TO_BYTE : BYTE
VAR_INPUT
    in : SINT;
END_VAR
    SINT_TO_BYTE := in;
END_FUNCTION

(********************
*
* Converts ULINT to LWORD
*
*********************)
FUNCTION ULINT_TO_LWORD : LWORD
VAR_INPUT
    in : ULINT;
END_VAR
    ULINT_TO_LWORD := in;
END_FUNCTION

(********************
*
* Converts ULINT to DWORD
*
*********************)
FUNCTION ULINT_TO_DWORD : DWORD
VAR_INPUT
    in : ULINT;
END_VAR
    ULINT_TO_DWORD := in;
END_FUNCTION

(********************
*
* Converts ULINT to WORD
*
*********************)
FUNCTION ULINT_TO_WORD : WORD
VAR_INPUT
    in : ULINT;
END_VAR
    ULINT_TO_WORD := in;
END_FUNCTION

(********************
*
* Converts ULINT to BYTE
*
*********************)
FUNCTION ULINT_TO_BYTE : BYTE
VAR_INPUT
    in : ULINT;
END_VAR
    ULINT_TO_BYTE := in;
END_FUNCTION

(********************
*
* Converts UDINT to LWORD
*
*********************)
FUNCTION UDINT_TO_LWORD : LWORD
VAR_INPUT
    in : UDINT;
END_VAR
    UDINT_TO_LWORD := in;
END_FUNCTION

(********************
*
* Converts UDINT to DWORD
*
*********************)
FUNCTION UDINT_TO_DWORD : DWORD
VAR_INPUT
    in : UDINT;
END_VAR
    UDINT_TO_DWORD := in;
END_FUNCTION

(********************
*
* Converts UDINT to WORD
*
*********************)
FUNCTION UDINT_TO_WORD : WORD
VAR_INPUT
    in : UDINT;
END_VAR
    UDINT_TO_WORD := in;
END_FUNCTION

(********************
*
* Converts UDINT to BYTE
*
*********************)
FUNCTION UDINT_TO_BYTE : BYTE
VAR_INPUT
    in : UDINT;
END_VAR
    UDINT_TO_BYTE := in;
END_FUNCTION

(********************
*
* Converts UINT to LWORD
*
*********************)
FUNCTION UINT_TO_LWORD : LWORD
VAR_INPUT
    in : UINT;
END_VAR
    UINT_TO_LWORD := in;
END_FUNCTION

(********************
*
* Converts UINT to DWORD
*
*********************)
FUNCTION UINT_TO_DWORD : DWORD
VAR_INPUT
    in : UINT;
END_VAR
    UINT_TO_DWORD := in;
END_FUNCTION

(********************
*
* Converts UINT to WORD
*
*********************)
FUNCTION UINT_TO_WORD : WORD
VAR_INPUT
    in : UINT;
END_VAR
    UINT_TO_WORD := in;
END_FUNCTION

(********************
*
* Converts UINT to BYTE
*
*********************)
FUNCTION UINT_TO_BYTE : BYTE
VAR_INPUT
    in : UINT;
END_VAR
    UINT_TO_BYTE := in;
END_FUNCTION

(********************
*
* Converts USINT to LWORD
*
*********************)
FUNCTION USINT_TO_LWORD : LWORD
VAR_INPUT
    in : USINT;
END_VAR
    USINT_TO_LWORD := in;
END_FUNCTION

(********************
*
* Converts USINT to DWORD
*
*********************)
FUNCTION USINT_TO_DWORD : DWORD
VAR_INPUT
    in : USINT;
END_VAR
    USINT_TO_DWORD := in;
END_FUNCTION

(********************
*
* Converts USINT to WORD
*
*********************)
FUNCTION USINT_TO_WORD : WORD
VAR_INPUT
    in : USINT;
END_VAR
    USINT_TO_WORD := in;
END_FUNCTION

(********************
*
* Converts USINT to BYTE
*
*********************)
FUNCTION USINT_TO_BYTE : BYTE
VAR_INPUT
    in : USINT;
END_VAR
    USINT_TO_BYTE := in;
END_FUNCTION

(* ---- bit_shift_functions.st ---- *)
(**************************
 *
 * ROL(IN, n)
 *
 * This operator implements a bitwise rotation of an operand to the left.
 * IN is shifted n-times to the left,
 * whereby the highest bit from the right is again inserted.
 *
*************************)
{external}
FUNCTION ROL<T : ANY_BIT> : T
VAR_INPUT
    IN : T;
    n : UDINT;
END_VAR
END_FUNCTION

(**************************
 *
 * ROR(IN, n)
 *
 * This operator implements a bitwise rotation of an operand to the right.
 * IN is shifted n-times to the right,
 * whereby the lowest bit from the left is again inserted.
 *
*************************)
{external}
FUNCTION ROR<T: ANY_BIT> : T
VAR_INPUT
    IN : T;
    n : UDINT;
END_VAR
END_FUNCTION

(* ---- date_time_conversion.st ---- *)
(********************
*
* Converts DT/LDT to DATE
*
*********************)
{external}
FUNCTION DATE_AND_TIME_TO_DATE : DATE
VAR_INPUT
    in : DT;
END_VAR
END_FUNCTION

(********************
*
* Converts DT/LDT to TOD/LTOD
*
*********************)
{external}
FUNCTION DATE_AND_TIME_TO_TIME_OF_DAY : TOD
VAR_INPUT
    in : DT;
END_VAR
END_FUNCTION

(********************
*
* Converts LTIME to TIME
*
*********************)
FUNCTION LTIME_TO_TIME : TIME
VAR_INPUT
    in : LTIME;
END_VAR
    LTIME_TO_TIME := in;
END_FUNCTION

(********************
*
* Converts TIME to LTIME
*
*********************)
FUNCTION TIME_TO_LTIME : LTIME
VAR_INPUT
    in : TIME;
END_VAR
    TIME_TO_LTIME := in;
END_FUNCTION

(********************
*
* Converts LDT to DT
*
*********************)
FUNCTION LDT_TO_DT : DT
VAR_INPUT
    in : LDT;
END_VAR
    LDT_TO_DT := in;
END_FUNCTION

(********************
*
* Converts LDT to DATE
*
*********************)
FUNCTION LDT_TO_DATE : DATE
VAR_INPUT
    in : LDT;
END_VAR
    LDT_TO_DATE := DATE_AND_TIME_TO_DATE(in);
END_FUNCTION

(********************
*
* Converts LDT to LTOD
*
*********************)
FUNCTION LDT_TO_LTOD : LTOD
VAR_INPUT
    in : LDT;
END_VAR
    LDT_TO_LTOD := DATE_AND_TIME_TO_TIME_OF_DAY(in);
END_FUNCTION

(********************
*
* Converts LDT to TOD
*
*********************)
FUNCTION LDT_TO_TOD : TOD
VAR_INPUT
    in : LDT;
END_VAR
    LDT_TO_TOD := DATE_AND_TIME_TO_TIME_OF_DAY(in);
END_FUNCTION

(********************
*
* Converts DT to LDT
*
*********************)
FUNCTION DT_TO_LDT : LDT
VAR_INPUT
    in : DT;
END_VAR
    DT_TO_LDT := in;
END_FUNCTION

(********************
*
* Converts DT to DATE
*
*********************)
FUNCTION DT_TO_DATE : DATE
VAR_INPUT
    in : DT;
END_VAR
    DT_TO_DATE := DATE_AND_TIME_TO_DATE(in);
END_FUNCTION

(********************
*
* Converts DT to LTOD
*
*********************)
FUNCTION DT_TO_LTOD : LTOD
VAR_INPUT
    in : DT;
END_VAR
    DT_TO_LTOD := DATE_AND_TIME_TO_TIME_OF_DAY(in);
END_FUNCTION

(********************
*
* Converts DT to TOD
*
*********************)
FUNCTION DT_TO_TOD : TOD
VAR_INPUT
    in : DT;
END_VAR
    DT_TO_TOD := DATE_AND_TIME_TO_TIME_OF_DAY(in);
END_FUNCTION

(********************
*
* Converts LTOD to TOD
*
*********************)
FUNCTION LTOD_TO_TOD : TOD
VAR_INPUT
    in : LTOD;
END_VAR
    LTOD_TO_TOD := in;
END_FUNCTION

(********************
*
* Converts TOD to LTOD
*
*********************)
FUNCTION TOD_TO_LTOD : LTOD
VAR_INPUT
    in : TOD;
END_VAR
    TOD_TO_LTOD := in;
END_FUNCTION

(* ---- date_time_extra_functions.st ---- *)
(********************
*
* Concatenates DATE and TOD to DT
*
*********************)
{external}
FUNCTION CONCAT_DATE_TOD : DT
VAR_INPUT
    date_input : DATE;
    tod_input : TOD;
END_VAR
END_FUNCTION

(********************
*
* Concatenates DATE and LTOD to DT
*
*********************)
FUNCTION CONCAT_DATE_LTOD : DT
VAR_INPUT
    date_input : DATE;
    tod_input : LTOD;
END_VAR
    CONCAT_DATE_LTOD := CONCAT_DATE_TOD(date_input, tod_input);
END_FUNCTION

(********************
*
* Concatenates year, month and day of type ANY_INT to DATE
*
*********************)
{external}
FUNCTION CONCAT_DATE <T: ANY_INT> : DATE
VAR_INPUT
    year : T;
    month : T;
    day : T;
END_VAR
END_FUNCTION

(********************
*
* Concatenates hour, minute, second, millisecond of type ANY_INT to TOD
*
*********************)
{external}
FUNCTION CONCAT_TOD <T: ANY_INT> : TOD
VAR_INPUT
    hour : T;
    minute : T;
    second : T;
    millisecond : T;
END_VAR
END_FUNCTION

(********************
*
* Concatenates hour, minute, second, millisecond of type ANY_INT to LTOD
*
*********************)
FUNCTION CONCAT_LTOD <T: ANY_INT> : LTOD
VAR_INPUT
    hour : T;
    minute : T;
    second : T;
    millisecond : T;
END_VAR
END_FUNCTION

(* Specialized implementation of CONCAT_LTOD for SINT *)
FUNCTION CONCAT_LTOD__SINT : LTOD
VAR_INPUT
    hour : SINT;
    minute : SINT;
    second : SINT;
    millisecond : SINT;
END_VAR
    CONCAT_LTOD__SINT := CONCAT_TOD(hour, minute, second, millisecond);
END_FUNCTION

(* Specialized implementation of CONCAT_LTOD for USINT *)
FUNCTION CONCAT_LTOD__USINT : LTOD
VAR_INPUT
    hour : USINT;
    minute : USINT;
    second : USINT;
    millisecond : USINT;
END_VAR
    CONCAT_LTOD__USINT := CONCAT_TOD(hour, minute, second, millisecond);
END_FUNCTION

(* Specialized implementation of CONCAT_LTOD for INT *)
FUNCTION CONCAT_LTOD__INT : LTOD
VAR_INPUT
    hour : INT;
    minute : INT;
    second : INT;
    millisecond : INT;
END_VAR
    CONCAT_LTOD__INT := CONCAT_TOD(hour, minute, second, millisecond);
END_FUNCTION

(* Specialized implementation of CONCAT_LTOD for UINT *)
FUNCTION CONCAT_LTOD__UINT : LTOD
VAR_INPUT
    hour : UINT;
    minute : UINT;
    second : UINT;
    millisecond : UINT;
END_VAR
    CONCAT_LTOD__UINT := CONCAT_TOD(hour, minute, second, millisecond);
END_FUNCTION

(* Specialized implementation of CONCAT_LTOD for DINT *)
FUNCTION CONCAT_LTOD__DINT : LTOD
VAR_INPUT
    hour : DINT;
    minute : DINT;
    second : DINT;
    millisecond : DINT;
END_VAR
    CONCAT_LTOD__DINT := CONCAT_TOD(hour, minute, second, millisecond);
END_FUNCTION

(* Specialized implementation of CONCAT_LTOD for UDINT *)
FUNCTION CONCAT_LTOD__UDINT : LTOD
VAR_INPUT
    hour : UDINT;
    minute : UDINT;
    second : UDINT;
    millisecond : UDINT;
END_VAR
    CONCAT_LTOD__UDINT := CONCAT_TOD(hour, minute, second, millisecond);
END_FUNCTION

(* Specialized implementation of CONCAT_LTOD for LINT *)
FUNCTION CONCAT_LTOD__LINT : LTOD
VAR_INPUT
    hour : LINT;
    minute : LINT;
    second : LINT;
    millisecond : LINT;
END_VAR
    CONCAT_LTOD__LINT := CONCAT_TOD(hour, minute, second, millisecond);
END_FUNCTION

(* Specialized implementation of CONCAT_LTOD for ULINT *)
FUNCTION CONCAT_LTOD__ULINT : LTOD
VAR_INPUT
    hour : ULINT;
    minute : ULINT;
    second : ULINT;
    millisecond : ULINT;
END_VAR
    CONCAT_LTOD__ULINT := CONCAT_TOD(hour, minute, second, millisecond);
END_FUNCTION

(********************
*
* Concatenates year, month, day, hour, minute, second, millisecond of type ANY_INT to DT
*
*********************)
FUNCTION CONCAT_DT <T: ANY_INT> : DT
VAR_INPUT
    year : T;
    month : T;
    day : T;
    hour : T;
    minute : T;
    second : T;
    millisecond : T;
END_VAR
END_FUNCTION

(* Specialized implementation of CONCAT_DT for INT *)
FUNCTION CONCAT_DT__INT : DT
VAR_INPUT
    year : INT;
    month : INT;
    day : INT;
    hour : INT;
    minute : INT;
    second : INT;
    millisecond : INT;
END_VAR
    CONCAT_DT__INT := CONCAT_DATE_TOD(CONCAT_DATE(year, month, day), CONCAT_TOD(hour, minute, second, millisecond));
END_FUNCTION

(* Specialized implementation of CONCAT_DT for UINT *)
FUNCTION CONCAT_DT__UINT : DT
VAR_INPUT
    year : UINT;
    month : UINT;
    day : UINT;
    hour : UINT;
    minute : UINT;
    second : UINT;
    millisecond : UINT;
END_VAR
    CONCAT_DT__UINT := CONCAT_DATE_TOD(CONCAT_DATE(year, month, day), CONCAT_TOD(hour, minute, second, millisecond));
END_FUNCTION

(* Specialized implementation of CONCAT_DT for DINT *)
FUNCTION CONCAT_DT__DINT : DT
VAR_INPUT
    year : DINT;
    month : DINT;
    day : DINT;
    hour : DINT;
    minute : DINT;
    second : DINT;
    millisecond : DINT;
END_VAR
    CONCAT_DT__DINT := CONCAT_DATE_TOD(CONCAT_DATE(year, month, day), CONCAT_TOD(hour, minute, second, millisecond));
END_FUNCTION

(* Specialized implementation of CONCAT_DT for UDINT *)
FUNCTION CONCAT_DT__UDINT : DT
VAR_INPUT
    year : UDINT;
    month : UDINT;
    day : UDINT;
    hour : UDINT;
    minute : UDINT;
    second : UDINT;
    millisecond : UDINT;
END_VAR
    CONCAT_DT__UDINT := CONCAT_DATE_TOD(CONCAT_DATE(year, month, day), CONCAT_TOD(hour, minute, second, millisecond));
END_FUNCTION

(* Specialized implementation of CONCAT_DT for LINT *)
FUNCTION CONCAT_DT__LINT : DT
VAR_INPUT
    year : LINT;
    month : LINT;
    day : LINT;
    hour : LINT;
    minute : LINT;
    second : LINT;
    millisecond : LINT;
END_VAR
    CONCAT_DT__LINT := CONCAT_DATE_TOD(CONCAT_DATE(year, month, day), CONCAT_TOD(hour, minute, second, millisecond));
END_FUNCTION

(* Specialized implementation of CONCAT_DT for ULINT *)
FUNCTION CONCAT_DT__ULINT : DT
VAR_INPUT
    year : ULINT;
    month : ULINT;
    day : ULINT;
    hour : ULINT;
    minute : ULINT;
    second : ULINT;
    millisecond : ULINT;
END_VAR
    CONCAT_DT__ULINT := CONCAT_DATE_TOD(CONCAT_DATE(year, month, day), CONCAT_TOD(hour, minute, second, millisecond));
END_FUNCTION

(********************
*
* Concatenates year, month, day, hour, minute, second, millisecond of type ANY_INT to LDT
*
*********************)
FUNCTION CONCAT_LDT <T: ANY_INT> : LDT
VAR_INPUT
    year : T;
    month : T;
    day : T;
    hour : T;
    minute : T;
    second : T;
    millisecond : T;
END_VAR
END_FUNCTION

(* Specialized implementation of CONCAT_LDT for INT *)
FUNCTION CONCAT_LDT__INT : LDT
VAR_INPUT
    year : INT;
    month : INT;
    day : INT;
    hour : INT;
    minute : INT;
    second : INT;
    millisecond : INT;
END_VAR
    CONCAT_LDT__INT := CONCAT_DATE_LTOD(CONCAT_DATE(year, month, day), CONCAT_LTOD(hour, minute, second, millisecond));
END_FUNCTION

(* Specialized implementation of CONCAT_LDT for UINT *)
FUNCTION CONCAT_LDT__UINT : LDT
VAR_INPUT
    year : UINT;
    month : UINT;
    day : UINT;
    hour : UINT;
    minute : UINT;
    second : UINT;
    millisecond : UINT;
END_VAR
    CONCAT_LDT__UINT := CONCAT_DATE_LTOD(CONCAT_DATE(year, month, day), CONCAT_LTOD(hour, minute, second, millisecond));
END_FUNCTION

(* Specialized implementation of CONCAT_LDT for DINT *)
FUNCTION CONCAT_LDT__DINT : LDT
VAR_INPUT
    year : DINT;
    month : DINT;
    day : DINT;
    hour : DINT;
    minute : DINT;
    second : DINT;
    millisecond : DINT;
END_VAR
    CONCAT_LDT__DINT := CONCAT_DATE_LTOD(CONCAT_DATE(year, month, day), CONCAT_LTOD(hour, minute, second, millisecond));
END_FUNCTION

(* Specialized implementation of CONCAT_LDT for UDINT *)
FUNCTION CONCAT_LDT__UDINT : LDT
VAR_INPUT
    year : UDINT;
    month : UDINT;
    day : UDINT;
    hour : UDINT;
    minute : UDINT;
    second : UDINT;
    millisecond : UDINT;
END_VAR
    CONCAT_LDT__UDINT := CONCAT_DATE_LTOD(CONCAT_DATE(year, month, day), CONCAT_LTOD(hour, minute, second, millisecond));
END_FUNCTION

(* Specialized implementation of CONCAT_LDT for LINT *)
FUNCTION CONCAT_LDT__LINT : LDT
VAR_INPUT
    year : LINT;
    month : LINT;
    day : LINT;
    hour : LINT;
    minute : LINT;
    second : LINT;
    millisecond : LINT;
END_VAR
    CONCAT_LDT__LINT := CONCAT_DATE_LTOD(CONCAT_DATE(year, month, day), CONCAT_LTOD(hour, minute, second, millisecond));
END_FUNCTION

(* Specialized implementation of CONCAT_LDT for ULINT *)
FUNCTION CONCAT_LDT__ULINT : LDT
VAR_INPUT
    year : ULINT;
    month : ULINT;
    day : ULINT;
    hour : ULINT;
    minute : ULINT;
    second : ULINT;
    millisecond : ULINT;
END_VAR
    CONCAT_LDT__ULINT := CONCAT_DATE_LTOD(CONCAT_DATE(year, month, day), CONCAT_LTOD(hour, minute, second, millisecond));
END_FUNCTION

(********************
*
* Splits DATE into year, month, day of type ANY_INT
*
*********************)
FUNCTION SPLIT_DATE <T: ANY_INT> : INT
VAR_INPUT
    in : DATE;
END_VAR
VAR_OUTPUT
    year : T;
    month : T;
    day : T;
END_VAR
END_FUNCTION

(* Specialized implementation of SPLIT_DATE for INT *)
{external}
FUNCTION SPLIT_DATE__INT : INT
VAR_INPUT
    in : DATE;
END_VAR
VAR_OUTPUT
    year : INT;
    month : INT;
    day : INT;
END_VAR
END_FUNCTION

(* Specialized implementation of SPLIT_DATE for UINT *)
{external}
FUNCTION SPLIT_DATE__UINT : INT
VAR_INPUT
    in : DATE;
END_VAR
VAR_OUTPUT
    year : UINT;
    month : UINT;
    day : UINT;
END_VAR
END_FUNCTION

(* Specialized implementation of SPLIT_DATE for DINT *)
{external}
FUNCTION SPLIT_DATE__DINT : INT
VAR_INPUT
    in : DATE;
END_VAR
VAR_OUTPUT
    year : DINT;
    month : DINT;
    day : DINT;
END_VAR
END_FUNCTION

(* Specialized implementation of SPLIT_DATE for UDINT *)
{external}
FUNCTION SPLIT_DATE__UDINT : INT
VAR_INPUT
    in : DATE;
END_VAR
VAR_OUTPUT
    year : UDINT;
    month : UDINT;
    day : UDINT;
END_VAR
END_FUNCTION

(* Specialized implementation of SPLIT_DATE for LINT *)
{external}
FUNCTION SPLIT_DATE__LINT : INT
VAR_INPUT
    in : DATE;
END_VAR
VAR_OUTPUT
    year : LINT;
    month : LINT;
    day : LINT;
END_VAR
END_FUNCTION

(* Specialized implementation of SPLIT_DATE for ULINT *)
{external}
FUNCTION SPLIT_DATE__ULINT : INT
VAR_INPUT
    in : DATE;
END_VAR
VAR_OUTPUT
    year : ULINT;
    month : ULINT;
    day : ULINT;
END_VAR
END_FUNCTION

(********************
*
* Splits TOD into hour, minute, second, millisecond of type ANY_INT
*
*********************)
FUNCTION SPLIT_TOD <T: ANY_INT> : INT
VAR_INPUT
    in : TOD;
END_VAR
VAR_OUTPUT
    hour : T;
    minute : T;
    second : T;
    millisecond : T;
END_VAR
END_FUNCTION

(* Specialized implementation of SPLIT_TOD for INT *)
{external}
FUNCTION SPLIT_TOD__INT : INT
VAR_INPUT
    in : TOD;
END_VAR
VAR_OUTPUT
    hour : INT;
    minute : INT;
    second : INT;
    millisecond : INT;
END_VAR
END_FUNCTION

(* Specialized implementation of SPLIT_TOD for UINT *)
{external}
FUNCTION SPLIT_TOD__UINT : INT
VAR_INPUT
    in : TOD;
END_VAR
VAR_OUTPUT
    hour : UINT;
    minute : UINT;
    second : UINT;
    millisecond : UINT;
END_VAR
END_FUNCTION

(* Specialized implementation of SPLIT_TOD for DINT *)
{external}
FUNCTION SPLIT_TOD__DINT : INT
VAR_INPUT
    in : TOD;
END_VAR
VAR_OUTPUT
    hour : DINT;
    minute : DINT;
    second : DINT;
    millisecond : DINT;
END_VAR
END_FUNCTION

(* Specialized implementation of SPLIT_TOD for UDINT *)
{external}
FUNCTION SPLIT_TOD__UDINT : INT
VAR_INPUT
    in : TOD;
END_VAR
VAR_OUTPUT
    hour : UDINT;
    minute : UDINT;
    second : UDINT;
    millisecond : UDINT;
END_VAR
END_FUNCTION

(* Specialized implementation of SPLIT_TOD for LINT *)
{external}
FUNCTION SPLIT_TOD__LINT : INT
VAR_INPUT
    in : TOD;
END_VAR
VAR_OUTPUT
    hour : LINT;
    minute : LINT;
    second : LINT;
    millisecond : LINT;
END_VAR
END_FUNCTION

(* Specialized implementation of SPLIT_TOD for ULINT *)
{external}
FUNCTION SPLIT_TOD__ULINT : INT
VAR_INPUT
    in : TOD;
END_VAR
VAR_OUTPUT
    hour : ULINT;
    minute : ULINT;
    second : ULINT;
    millisecond : ULINT;
END_VAR
END_FUNCTION

(********************
*
* Splits LTOD into hour, minute, second, millisecond of type ANY_INT
*
*********************)
FUNCTION SPLIT_LTOD <T: ANY_INT> : INT
VAR_INPUT
    in : LTOD;
END_VAR
VAR_OUTPUT
    hour : T;
    minute : T;
    second : T;
    millisecond : T;
END_VAR
END_FUNCTION

(* Specialized implementation of SPLIT_LTOD for INT *)
FUNCTION SPLIT_LTOD__INT : INT
VAR_INPUT
    in : LTOD;
END_VAR
VAR_OUTPUT
    hour : INT;
    minute : INT;
    second : INT;
    millisecond : INT;
END_VAR
    SPLIT_LTOD__INT := SPLIT_TOD__INT(in, hour, minute, second, millisecond);
END_FUNCTION

(* Specialized implementation of SPLIT_LTOD for UINT *)
FUNCTION SPLIT_LTOD__UINT : INT
VAR_INPUT
    in : LTOD;
END_VAR
VAR_OUTPUT
    hour : UINT;
    minute : UINT;
    second : UINT;
    millisecond : UINT;
END_VAR
    SPLIT_LTOD__UINT := SPLIT_TOD__UINT(in, hour, minute, second, millisecond);
END_FUNCTION

(* Specialized implementation of SPLIT_LTOD for DINT *)
FUNCTION SPLIT_LTOD__DINT : INT
VAR_INPUT
    in : LTOD;
END_VAR
VAR_OUTPUT
    hour : DINT;
    minute : DINT;
    second : DINT;
    millisecond : DINT;
END_VAR
    SPLIT_LTOD__DINT := SPLIT_TOD__DINT(in, hour, minute, second, millisecond);
END_FUNCTION

(* Specialized implementation of SPLIT_LTOD for UDINT *)
FUNCTION SPLIT_LTOD__UDINT : INT
VAR_INPUT
    in : LTOD;
END_VAR
VAR_OUTPUT
    hour : UDINT;
    minute : UDINT;
    second : UDINT;
    millisecond : UDINT;
END_VAR
    SPLIT_LTOD__UDINT := SPLIT_TOD__UDINT(in, hour, minute, second, millisecond);
END_FUNCTION

(* Specialized implementation of SPLIT_LTOD for LINT *)
FUNCTION SPLIT_LTOD__LINT : INT
VAR_INPUT
    in : LTOD;
END_VAR
VAR_OUTPUT
    hour : LINT;
    minute : LINT;
    second : LINT;
    millisecond : LINT;
END_VAR
    SPLIT_LTOD__LINT := SPLIT_TOD__LINT(in, hour, minute, second, millisecond);
END_FUNCTION

(* Specialized implementation of SPLIT_LTOD for ULINT *)
FUNCTION SPLIT_LTOD__ULINT : INT
VAR_INPUT
    in : LTOD;
END_VAR
VAR_OUTPUT
    hour : ULINT;
    minute : ULINT;
    second : ULINT;
    millisecond : ULINT;
END_VAR
    SPLIT_LTOD__ULINT := SPLIT_TOD__ULINT(in, hour, minute, second, millisecond);
END_FUNCTION

(********************
*
* Splits DT into year, month, day, hour, minute, second, millisecond of type ANY_INT
*
*********************)
FUNCTION SPLIT_DT <T: ANY_INT> : INT
VAR_INPUT
    in : DT;
END_VAR
VAR_OUTPUT
    year : T;
    month : T;
    day : T;
    hour : T;
    minute : T;
    second : T;
    millisecond : T;
END_VAR
END_FUNCTION

(* Specialized implementation of SPLIT_DT for INT *)
{external}
FUNCTION SPLIT_DT__INT : INT
VAR_INPUT
    in : DT;
END_VAR
VAR_OUTPUT
    year : INT;
    month : INT;
    day : INT;
    hour : INT;
    minute : INT;
    second : INT;
    millisecond : INT;
END_VAR
END_FUNCTION

(* Specialized implementation of SPLIT_DT for UINT *)
{external}
FUNCTION SPLIT_DT__UINT : INT
VAR_INPUT
    in : DT;
END_VAR
VAR_OUTPUT
    year : UINT;
    month : UINT;
    day : UINT;
    hour : UINT;
    minute : UINT;
    second : UINT;
    millisecond : UINT;
END_VAR
END_FUNCTION

(* Specialized implementation of SPLIT_DT for DINT *)
{external}
FUNCTION SPLIT_DT__DINT : INT
VAR_INPUT
    in : DT;
END_VAR
VAR_OUTPUT
    year : DINT;
    month : DINT;
    day : DINT;
    hour : DINT;
    minute : DINT;
    second : DINT;
    millisecond : DINT;
END_VAR
END_FUNCTION

(* Specialized implementation of SPLIT_DT for UDINT *)
{external}
FUNCTION SPLIT_DT__UDINT : INT
VAR_INPUT
    in : DT;
END_VAR
VAR_OUTPUT
    year : UDINT;
    month : UDINT;
    day : UDINT;
    hour : UDINT;
    minute : UDINT;
    second : UDINT;
    millisecond : UDINT;
END_VAR
END_FUNCTION

(* Specialized implementation of SPLIT_DT for LINT *)
{external}
FUNCTION SPLIT_DT__LINT : INT
VAR_INPUT
    in : DT;
END_VAR
VAR_OUTPUT
    year : LINT;
    month : LINT;
    day : LINT;
    hour : LINT;
    minute : LINT;
    second : LINT;
    millisecond : LINT;
END_VAR
END_FUNCTION

(* Specialized implementation of SPLIT_DT for ULINT *)
{external}
FUNCTION SPLIT_DT__ULINT : INT
VAR_INPUT
    in : DT;
END_VAR
VAR_OUTPUT
    year : ULINT;
    month : ULINT;
    day : ULINT;
    hour : ULINT;
    minute : ULINT;
    second : ULINT;
    millisecond : ULINT;
END_VAR
END_FUNCTION

(********************
*
* Splits LDT into year, month, day, hour, minute, second, millisecond of type ANY_INT
*
*********************)
FUNCTION SPLIT_LDT <T: ANY_INT> : INT
VAR_INPUT
    in : LDT;
END_VAR
VAR_OUTPUT
    year : T;
    month : T;
    day : T;
    hour : T;
    minute : T;
    second : T;
    millisecond : T;
END_VAR
END_FUNCTION

(* Specialized implementation of SPLIT_LDT for INT *)
{external}
FUNCTION SPLIT_LDT__INT : INT
VAR_INPUT
    in : LDT;
END_VAR
VAR_OUTPUT
    year : INT;
    month : INT;
    day : INT;
    hour : INT;
    minute : INT;
    second : INT;
    millisecond : INT;
END_VAR
    SPLIT_LDT__INT := SPLIT_DT__INT(in, year, month, day, hour, minute, second, millisecond);
END_FUNCTION

(* Specialized implementation of SPLIT_LDT for UINT *)
{external}
FUNCTION SPLIT_LDT__UINT : INT
VAR_INPUT
    in : LDT;
END_VAR
VAR_OUTPUT
    year : UINT;
    month : UINT;
    day : UINT;
    hour : UINT;
    minute : UINT;
    second : UINT;
    millisecond : UINT;
END_VAR
    SPLIT_LDT__UINT := SPLIT_DT__UINT(in, year, month, day, hour, minute, second, millisecond);
END_FUNCTION

(* Specialized implementation of SPLIT_LDT for DINT *)
{external}
FUNCTION SPLIT_LDT__DINT : INT
VAR_INPUT
    in : LDT;
END_VAR
VAR_OUTPUT
    year : DINT;
    month : DINT;
    day : DINT;
    hour : DINT;
    minute : DINT;
    second : DINT;
    millisecond : DINT;
END_VAR
    SPLIT_LDT__DINT := SPLIT_DT__DINT(in, year, month, day, hour, minute, second, millisecond);
END_FUNCTION

(* Specialized implementation of SPLIT_LDT for UDINT *)
{external}
FUNCTION SPLIT_LDT__UDINT : INT
VAR_INPUT
    in : LDT;
END_VAR
VAR_OUTPUT
    year : UDINT;
    month : UDINT;
    day : UDINT;
    hour : UDINT;
    minute : UDINT;
    second : UDINT;
    millisecond : UDINT;
END_VAR
    SPLIT_LDT__UDINT := SPLIT_DT__UDINT(in, year, month, day, hour, minute, second, millisecond);
END_FUNCTION

(* Specialized implementation of SPLIT_LDT for LINT *)
{external}
FUNCTION SPLIT_LDT__LINT : INT
VAR_INPUT
    in : LDT;
END_VAR
VAR_OUTPUT
    year : LINT;
    month : LINT;
    day : LINT;
    hour : LINT;
    minute : LINT;
    second : LINT;
    millisecond : LINT;
END_VAR
    SPLIT_LDT__LINT := SPLIT_DT__LINT(in, year, month, day, hour, minute, second, millisecond);
END_FUNCTION

(* Specialized implementation of SPLIT_LDT for ULINT *)
{external}
FUNCTION SPLIT_LDT__ULINT : INT
VAR_INPUT
    in : LDT;
END_VAR
VAR_OUTPUT
    year : ULINT;
    month : ULINT;
    day : ULINT;
    hour : ULINT;
    minute : ULINT;
    second : ULINT;
    millisecond : ULINT;
END_VAR
    SPLIT_LDT__ULINT := SPLIT_DT__ULINT(in, year, month, day, hour, minute, second, millisecond);
END_FUNCTION

(********************
*
* Returns day of week form given DATE in SINT
* 0 -> sunday, 1 -> monday, ..., 6 -> saturday
*
*********************)
{external}
FUNCTION DAY_OF_WEEK : SINT
VAR_INPUT
    in : DATE;
END_VAR
END_FUNCTION

(* ---- date_time_numeric_functions.st ---- *)
(* Specialized implementation of ADD for TIME *)
FUNCTION ADD__TIME__TIME: TIME
VAR_INPUT
    IN1: TIME;
    IN2: TIME;
END_VAR
    ADD__TIME__TIME := ADD_TIME(IN1, IN2);
END_FUNCTION

(********************
*
* This operator returns the value of adding up two TIME operands.
*
*********************)
{external}
FUNCTION ADD_TIME: TIME
VAR_INPUT
    IN1: TIME;
    IN2: TIME;
END_VAR
END_FUNCTION

(********************
*
* This operator returns the value of adding up two LTIME operands.
*
*********************)
FUNCTION ADD_LTIME: LTIME
VAR_INPUT
    IN1: LTIME;
    IN2: LTIME;
END_VAR
    ADD_LTIME := ADD_TIME(IN1, IN2);
END_FUNCTION

(* Specialized implementation of ADD for TOD *)
FUNCTION ADD__TIME_OF_DAY__TIME: TOD
VAR_INPUT
    IN1: TOD;
    IN2: TIME;
END_VAR
    ADD__TIME_OF_DAY__TIME := ADD_TOD_TIME(IN1, IN2);
END_FUNCTION

(********************
*
* This operator returns the value of adding up TOD and TIME.
* Panic on overflow
*
*********************)
{external}
FUNCTION ADD_TOD_TIME: TOD
VAR_INPUT
    IN1: TOD;
    IN2: TIME;
END_VAR
END_FUNCTION

(********************
*
* This operator returns the value of adding up LTOD and LTIME.
* Panic on overflow
*
*********************)
FUNCTION ADD_LTOD_LTIME: LTOD
VAR_INPUT
    IN1: LTOD;
    IN2: LTIME;
END_VAR
    ADD_LTOD_LTIME := ADD_TOD_TIME(IN1, IN2);
END_FUNCTION

(* Specialized implementation of ADD for DT *)
FUNCTION ADD__DATE_AND_TIME__TIME: DT
VAR_INPUT
    IN1: DT;
    IN2: TIME;
END_VAR
    ADD__DATE_AND_TIME__TIME := ADD_DT_TIME(IN1, IN2);
END_FUNCTION

(********************
*
* This operator returns the value of adding up DT and TIME.
* Panic on overflow
*
*********************)
{external}
FUNCTION ADD_DT_TIME: DT
VAR_INPUT
    IN1: DT;
    IN2: TIME;
END_VAR
END_FUNCTION

(********************
*
* This operator returns the value of adding up LDT and LTIME.
* Panic on overflow
*
*********************)
FUNCTION ADD_LDT_LTIME: LDT
VAR_INPUT
    IN1: LDT;
    IN2: LTIME;
END_VAR
    ADD_LDT_LTIME := ADD_DT_TIME(IN1, IN2);
END_FUNCTION

(* Specialized implementation of SUB for TIME *)
FUNCTION SUB__TIME__TIME: TIME
VAR_INPUT
    IN1: TIME;
    IN2: TIME;
END_VAR
    SUB__TIME__TIME := SUB_TIME(IN1, IN2);
END_FUNCTION

(********************
*
* This operator produces the subtraction of two TIME operands
*
*********************)
{external}
FUNCTION SUB_TIME: TIME
VAR_INPUT
    IN1: TIME;
    IN2: TIME;
END_VAR
END_FUNCTION

(********************
*
* This operator produces the subtraction of two LTIME operands
*
*********************)
FUNCTION SUB_LTIME: LTIME
VAR_INPUT
    IN1: LTIME;
    IN2: LTIME;
END_VAR
    SUB_LTIME := SUB_TIME(IN1, IN2);
END_FUNCTION

(* Specialized implementation of SUB for DATE *)
FUNCTION SUB__DATE__DATE: TIME
VAR_INPUT
    IN1: DATE;
    IN2: DATE;
END_VAR
    SUB__DATE__DATE := SUB_DATE_DATE(IN1, IN2);
END_FUNCTION

(********************
*
* This operator produces the subtraction of two DATE operands returning TIME
* Panic on overflow
*
*********************)
{external}
FUNCTION SUB_DATE_DATE: TIME
VAR_INPUT
    IN1: DATE;
    IN2: DATE;
END_VAR
END_FUNCTION

(********************
*
* This operator produces the subtraction of two LDATE operands returning LTIME
* Panic on overflow
*
*********************)
FUNCTION SUB_LDATE_LDATE: LTIME
VAR_INPUT
    IN1: LDATE;
    IN2: LDATE;
END_VAR
    SUB_LDATE_LDATE := SUB_DATE_DATE(IN1, IN2);
END_FUNCTION

(* Specialized implementation of SUB for TOD and TIME *)
FUNCTION SUB__TIME_OF_DAY__TIME: TOD
VAR_INPUT
    IN1: TOD;
    IN2: TIME;
END_VAR
    SUB__TIME_OF_DAY__TIME := SUB_TOD_TIME(IN1, IN2);
END_FUNCTION

(********************
*
* This operator produces the subtraction of TOD and TIME returning TOD
* Panic on overflow
*
*********************)
{external}
FUNCTION SUB_TOD_TIME: TOD
VAR_INPUT
    IN1: TOD;
    IN2: TIME;
END_VAR
END_FUNCTION

(********************
*
* This operator produces the subtraction of LTOD and LTIME returning LTOD
* Panic on overflow
*
*********************)
FUNCTION SUB_LTOD_LTIME: LTOD
VAR_INPUT
    IN1: LTOD;
    IN2: LTIME;
END_VAR
    SUB_LTOD_LTIME := SUB_TOD_TIME(IN1, IN2);
END_FUNCTION

(* Specialized implementation of SUB for TOD *)
FUNCTION SUB__TIME_OF_DAY__TIME_OF_DAY: TIME
VAR_INPUT
    IN1: TOD;
    IN2: TOD;
END_VAR
    SUB__TIME_OF_DAY__TIME_OF_DAY := SUB_TOD_TOD(IN1, IN2);
END_FUNCTION

(********************
*
* This operator produces the subtraction of two TOD operands returning TIME
* Panic on overflow
*
*********************)
{external}
FUNCTION SUB_TOD_TOD: TIME
VAR_INPUT
    IN1: TOD;
    IN2: TOD;
END_VAR
END_FUNCTION

(********************
*
* This operator produces the subtraction of two LTOD operands returning LTIME
* Panic on overflow
*
*********************)
FUNCTION SUB_LTOD_LTOD: LTIME
VAR_INPUT
    IN1: LTOD;
    IN2: LTOD;
END_VAR
    SUB_LTOD_LTOD := SUB_TOD_TOD(IN1, IN2);
END_FUNCTION

(* Specialized implementation of SUB for DT and TIME *)
FUNCTION SUB__DATE_AND_TIME__TIME: DT
VAR_INPUT
    IN1: DT;
    IN2: TIME;
END_VAR
    SUB__DATE_AND_TIME__TIME := SUB_DT_TIME(IN1, IN2);
END_FUNCTION

(********************
*
* This operator produces the subtraction of DT and TIME returning DT
* Panic on overflow
*
*********************)
{external}
FUNCTION SUB_DT_TIME: DT
VAR_INPUT
    IN1: DT;
    IN2: TIME;
END_VAR
END_FUNCTION

(********************
*
* This operator produces the subtraction of LDT and LTIME returning LDT
* Panic on overflow
*
*********************)
FUNCTION SUB_LDT_LTIME: LDT
VAR_INPUT
    IN1: LDT;
    IN2: LTIME;
END_VAR
    SUB_LDT_LTIME := SUB_DT_TIME(IN1, IN2);
END_FUNCTION

(* Specialized implementation of SUB for DT *)
FUNCTION SUB__DATE_AND_TIME__DATE_AND_TIME: TIME
VAR_INPUT
    IN1: DT;
    IN2: DT;
END_VAR
    SUB__DATE_AND_TIME__DATE_AND_TIME := SUB_DT_DT(IN1, IN2);
END_FUNCTION

(********************
*
* This operator produces the subtraction of two DT operands returning TIME
* Panic on overflow
*
*********************)
{external}
FUNCTION SUB_DT_DT: TIME
VAR_INPUT
    IN1: DT;
    IN2: DT;
END_VAR
END_FUNCTION

(********************
*
* This operator produces the subtraction of two LDT operands returning LTIME
* Panic on overflow
*
*********************)
FUNCTION SUB_LDT_LDT: LTIME
VAR_INPUT
    IN1: LDT;
    IN2: LDT;
END_VAR
    SUB_LDT_LDT := SUB_DT_DT(IN1, IN2);
END_FUNCTION

(********************
*
* This operator produces the multiplication of TIME and ANY_NUM.
*
*********************)
FUNCTION MUL_TIME < T: ANY_NUM >: TIME
VAR_INPUT
    IN1: TIME;
    IN2: T;
END_VAR
END_FUNCTION

(********************
*
* This operator produces the multiplication of LTIME and ANY_NUM.
*
*********************)
FUNCTION MUL_LTIME < T: ANY_NUM >: LTIME
VAR_INPUT
    IN1: LTIME;
    IN2: T;
END_VAR
END_FUNCTION

(********************
*
* This operator produces the division of TIME and ANY_NUM.
*
*********************)
FUNCTION DIV_TIME < T: ANY_NUM >: TIME
VAR_INPUT
    IN1: TIME;
    IN2: T;
END_VAR
END_FUNCTION

(********************
*
* This operator produces the division of LTIME and ANY_NUM.
*
*********************)
FUNCTION DIV_LTIME < T: ANY_NUM >: LTIME
VAR_INPUT
    IN1: LTIME;
    IN2: T;
END_VAR
END_FUNCTION

(* ---- endianness_conversion_functions.st ---- *)
(******************************************************************************
Description: Converts data to big endian format from native endian format.
Input:
  - in: The input value in native endian format.
Return: The value converted to big endian format.
******************************************************************************)
{external}
FUNCTION TO_BIG_ENDIAN<T: ANY> : T
VAR_INPUT
    in : T;
END_VAR
END_FUNCTION

(******************************************************************************
Description: Converts data to little endian format from big endian format.
Input:
  - in: The input value in native endian format.
Return: The value converted to little endian format.
******************************************************************************)
{external}
FUNCTION TO_LITTLE_ENDIAN<T: ANY> : T
VAR_INPUT
    in : T;
END_VAR
END_FUNCTION

(******************************************************************************
Description: Converts data from big endian format to native endian format.
Input:
  - in: The input value in big endian format.
Return: The value converted to native endian format.
******************************************************************************)
{external}
FUNCTION FROM_BIG_ENDIAN<T: ANY> : T
VAR_INPUT
    in : T;
END_VAR
END_FUNCTION

(******************************************************************************
Description: Converts data from little endian format to native endian format.
Input:
  - in: The input value in little endian format.
Return: The value converted to native endian format.
******************************************************************************)
{external}
FUNCTION FROM_LITTLE_ENDIAN<T: ANY> : T
VAR_INPUT
    in : T;
END_VAR
END_FUNCTION
